// TIA Portal V20 export
TYPE "AZ_Struct_Drv2PLC"
   STRUCT
      RemoteIO_OUT : Word;
      OperNumSel_R : Word;
      FixedIO_OUT { S7_SetPoint := 'True'} : "AZ_FixedIO_Drv2PLC";
      PresentAlm : Word;
      DetectPos : DInt;
      DetectVel : DInt;
      CmdPos : DInt;
      Torque : Int;
      OpeCrnt : UInt;
      Information : DWord;
      Reserve : Word;
      ReadPrmID_R : Word;
      RW_Status : Word;
      WritePrmID_R : Word;
      ReadData : DInt;
      Monitor0 : DInt;
      Monitor1 : DInt;
      Monitor2 : DInt;
      Monitor3 : DInt;
   END_STRUCT;
END_TYPE
